(* IEC 61131-3 sources: sis-interlock-demo/pytests/golden/mini/tests/GVLs/Generated, 1 file *)

(* ---- GVL_TestsGenerated.gvl.st ---- *)
// AUTO-GENERATED by cemgen 1.0.0 — не редактировать: правьте матрицу и запустите
//   python -m cemgen generate <файл матрицы .csv или .xlsx>
// Матрица: TEST-U301-CEM, объект U-301, ревизия 1 от 2026-10-16, SHA-256 сетки 9067fda96ae55e67
// Назначение: экземпляры сгенерированных наборов coUnit: таблицы истинности голосования и сценарии
//             по матрице. {attribute 'linkalways'} обязателен: без него CODESYS выбрасывает GVL, на
//             которую никто не ссылается, и наборы молча пропадают.
// Автор:      pytest; код — генератор cemgen
// Версия:     1.0.0
// Документ:   docs/DESIGN.md, раздел «10. Генератор cemgen»; docs/cause_effect_matrix.md
// ВНИМАНИЕ:   код демонстрационный и не предназначен для систем безопасности. Реальная ПАЗ требует
//             определения SIL, сертифицированных аппаратных и программных средств и валидации по
//             ГОСТ Р МЭК 61511.
{attribute 'qualified_only'}
{attribute 'linkalways'}
VAR_GLOBAL
    fbVoteTruthTest : FB_VoteTruth_Test;   // таблицы истинности голосования (36 тестов)
    fbCemGen01Test  : FB_CemGen01_Test;    // сценарии по матрице, тесты 1–24
END_VAR
